Staubli VAL3: data.pjx

--- data.pjx ---
Parameters version=s8.10.3cs9_BS2093 stackSize=20000 millimeterUnit=true
Program file=start.pgx
Program file=stop.pgx
Data file=data.dtx

--- data.dtx ---
public frame fFrame[10]
  [0] = {fatherId=world[0]}
  [1] = {fatherId=world[0]}
  [2] = {fatherId=world[0]}
  [3] = {fatherId=world[0]}
  [4] = {fatherId=world[0]}
  [5] = {fatherId=world[0]}
  [6] = {fatherId=world[0]}
  [7] = {fatherId=world[0]}
  [8] = {fatherId=world[0]}
  [9] = {fatherId=world[0]}
public jointRx jHome = {j1=2.180132, j2=-34.106359, j3=121.0461159, j4=-3.0709494, j5=46.658106, j6=2.441583}
public mdesc mMdesc[40]
public pointRx pPointRx[30]
  [0] = {x=617.494944, y=437.693102, z=144.0206459, rx=0.508772, ry=175.411265, rz=0.199171, fatherId=world[0]}
  [1] = {x=617.494811, y=-390.105125, z=144.0205963, rx=0.508128, ry=175.410572, rz=0.199501, fatherId=world[0]}
  [2] = {fatherId=world[0]}
  [3] = {fatherId=world[0]}
  [4] = {fatherId=world[0]}
  [5] = {fatherId=world[0]}
  [6] = {fatherId=world[0]}
  [7] = {fatherId=world[0]}
  [8] = {fatherId=world[0]}
  [9] = {fatherId=world[0]}
  [10] = {fatherId=world[0]}
  [11] = {fatherId=world[0]}
  [12] = {fatherId=world[0]}
  [13] = {fatherId=world[0]}
  [14] = {fatherId=world[0]}
  [15] = {fatherId=world[0]}
  [16] = {fatherId=world[0]}
  [17] = {fatherId=world[0]}
  [18] = {fatherId=world[0]}
  [19] = {fatherId=world[0]}
  [20] = {fatherId=world[0]}
  [21] = {fatherId=world[0]}
  [22] = {fatherId=world[0]}
  [23] = {fatherId=world[0]}
  [24] = {fatherId=world[0]}
  [25] = {fatherId=world[0]}
  [26] = {fatherId=world[0]}
  [27] = {fatherId=world[0]}
  [28] = {fatherId=world[0]}
  [29] = {fatherId=world[0]}
public tool tTool[10]
  [0] = {fatherId=flange[0]}
  [1] = {fatherId=flange[0]}
  [2] = {fatherId=flange[0]}
  [3] = {fatherId=flange[0]}
  [4] = {fatherId=flange[0]}
  [5] = {fatherId=flange[0]}
  [6] = {fatherId=flange[0]}
  [7] = {fatherId=flange[0]}
  [8] = {fatherId=flange[0]}
  [9] = {fatherId=flange[0]}

--- start.pgx ---
program start()
begin
end

--- stop.pgx ---
program stop()
begin
end
